DATA_BLOCK "GDB_GRAPH_PressDemoAutoLoadPosition"
{ S7_Optimized_Access := 'TRUE' }
VERSION : 0.1
NON_RETAIN
"FB_GRAPH_PressDemoLoadPosition"
BEGIN
END_DATA_BLOCK
